FUNCTION_BLOCK FB_FourAxisTrajectory
// 四轴整表轨迹：上位机预检后下发 LREAL 位置点，本块收齐后统一执行。
// 正常流程：0 登记各段 -> 全部下发后 5 统一拼表 -> 0 就绪 -> 10 启动检查 -> 15 首点定位
//           -> 20 开外部给定 -> 30 取点 -> 40 保持末点 -> 60 关闭 -> 70 确认静止 -> 0。
// 异常流程：运动阶段转 50 减速，再经 40/60/70 退出，最后在 90 等待复位。
// 本块每 2 ms 调用一次；使能、点动、回原等基础控制在 FB_AxisControl 中。
// xGroupBusy 占用控制防止两块同时运动，但不能代替设备安全回路。
VAR_INPUT
    xAxesReady : BOOL; // 四轴已使能、回零、静止，供启动和首点定位完成时检查。
    xAbort : BOOL; // 外部联停：许可撤销、撤使能、停止、限位或手动命令冲突。
    nAbortReason : UINT; // MAIN 提供的首个联停原因，0 表示本扫描无联停。
    xAxisFault : BOOL; // 任一轴错误或 NC I/O 反馈无效，拒绝启动或触发联停。
END_VAR
VAR_IN_OUT
    Axes : ARRAY[1..4] OF AXIS_REF; // MAIN 传入的原始轴引用，VAR_IN_OUT 直接操作各 NC 轴接口。
END_VAR
VAR
    // 完整四轴位置表，只由本块分段写入；运行中不再接收上传。
    aPosition : ARRAY[1..4, 0..2099999] OF LREAL; // [轴号, 完整表点号]，所有点号从 0 开始，单位由 NC 配置决定。
    aConfig : ARRAY[1..4] OF ST_AxisConfig; // 启动时锁存参数，首点定位、运行及本次停车使用相同参数。
    aSet : ARRAY[1..4] OF ST_TrajectoryPoint; // 本周期四轴的位置、内部速度和加速度；内部速度用于减速停车。
    aEnable : ARRAY[1..4] OF MC_ExtSetPointGenEnable; // 四个外部给定开启实例；异步执行，等待 NC Enabled 反馈。
    aDisable : ARRAY[1..4] OF MC_ExtSetPointGenDisable; // 四个关闭实例；确认全部退出之前不交回手动。
    aMoveInit : ARRAY[1..4] OF MC_MoveAbsolute; // 四轴各自定位到轨迹首点，全部完成才同步执行位置表。
    aStopInit : ARRAY[1..4] OF MC_Stop; // 外部给定尚未开启时的停车，如取消首点定位。
    rtUpload : R_TRIG; // 本段四轴数据写完后的登记请求上升沿。
    rtAssemble : R_TRIG; // 全部段登记后的独立拼表请求上升沿，不自动启动运动。
    rtClear : R_TRIG; // 清除旧表计数和就绪状态的请求上升沿。
    rtStart : R_TRIG; // 完整位置表就绪后启动轨迹的请求上升沿。
    rtReset : R_TRIG; // 轨迹组故障复位请求上升沿，不复位各 NC 轴故障。
    tmHeartbeat : TON; // 上位机运行心跳超时定时器，启动检查/运动期间 1 秒不变则联停。
    tmEnable : TON; // 四轴外部给定开启阶段超时定时器，限时 5 秒。
    tmMoveInit : TON; // 四轴首点定位阶段超时定时器，限时 60 秒。
    tmExit : TON; // 关闭外部给定及确认退出阶段的超时定时器，限时 5 秒。
    udiLastHeartbeat : UDINT; // 上一扫描上位机运行心跳值，用于检测是否发生变化。
    udiSequence : UDINT; // 当前接收/执行位置表锁存的非零上传序号。
    nCount : UDINT; // 当前整条位置表锁存的单轴总点数，四根轴点数相同。
    nReceived : UDINT; // 已登记的单轴点数，表示段确认进度，不代表已拼入执行表。
    nLoaded : UDINT; // 四轴均已成功拼入执行表的点数。
    nSegment : UDINT; // 当前拼表源段号，从 0 开始，范围 0～20。
    nSegmentPoint : UDINT; // 当前源段内的起始点号，从 0 开始。
    nCopyCount : UDINT; // 本扫描每轴复制点数，受批次、段尾和总表尾三重限制。
    nCopyBytes : UDINT; // 本扫描每轴复制的字节数，等于点数乘 LREAL 大小。
    nSendPoint : UDINT; // 当前轨迹执行取点号，从 0 开始，不是实际到位点号。
    nPrevious : UDINT; // 差分计算前一点索引，首点处夹紧到有效表范围。
    nNext : UDINT; // 差分计算后一点索引，末点处夹紧到有效表范围。
    nHoldCycles : UINT; // 末点静止给定的保持扫描次数，每扫描为 2 ms。
    nStopCycles : UINT; // 减速阶段扫描计数，用于满足该阶段的最少扫描次数。
    nState : UINT; // 轨迹阶段码，数值与上位机监控和故障诊断一致。
    i : INT; // 四轴循环索引，范围 1～4。
    xAllEnabled : BOOL; // 四轴 NC 外部给定均已开启；不是四轴伺服使能汇总。
    xAllDisabled : BOOL; // 四轴外部给定均已关闭，相关开启、关闭和首点停止块均释放 Busy。
    xAllStopped : BOOL; // 四轴 NC 均未处于 Moving 状态；仅为本块此项汇总条件。
    xAllInitDone : BOOL; // 四个首点绝对定位块均输出 Done。
    xMovesIdle : BOOL; // 四个首点定位块均已释放 Busy。
    xEnablePending : BOOL; // 至少一个外部给定开启块仍忙，退出时先等待开启请求结束。
    xFeed : BOOL; // 本扫描需要向四轴发送外部位置给定。
    xValid : BOOL; // 当前轴配置、首点到位或内存复制批次的临时检查结果，每次检查重新赋值。
    xCommandAllowed : BOOL; // 轨迹命令来源为当前有效持有站，且本扫描未发生控制权交接。
    xStopCommand : BOOL; // 当前持有站发出的有效组停止保持命令。
    xUploadRequest : BOOL; // 本扫描获准处理的段登记请求；原始沿已消费后再过滤权限。
    xAssembleRequest : BOOL; // 本扫描获准处理的整表拼接请求。
    xClearRequest : BOOL; // 本扫描获准处理的清表请求。
    xStartRequest : BOOL; // 本扫描获准处理的轨迹启动请求。
    xResetRequest : BOOL; // 本扫描获准处理的轨迹组故障复位请求。
    xNormalStop : BOOL; // 正常人工停止，不作为 1007 故障。
    lrNewVelocity : LREAL; // 当前减速计算的下一扫描速度，单位为 NC 位置单位/秒。
    nBlockAxis : UINT; // 本扫描首个定位/开启块错误的轴，四轴循环结束后统一联停。
    nBlockSource : UINT; // 10=首点定位，11=开启外部给定。
    udiBlockError : UDINT; // 本扫描首个定位/开启块原始错误码，后续轴不能覆盖。
END_VAR
VAR CONSTANT
    // 保留原阶段数值及顺序，供监控和原有区间判断使用。
    cStateIdle : UINT := 0; // 空闲及收段。
    cStateAssemble : UINT := 5; // 拼接已确认的点位段。
    cStateCheckStart : UINT := 10; // 检查轴配置和启动条件。
    cStateMoveToFirstPoint : UINT := 15; // 四轴定位到首点。
    cStateEnableSetpoint : UINT := 20; // 开启外部给定。
    cStateRun : UINT := 30; // 按 2 ms 送点。
    cStateHoldLastPoint : UINT := 40; // 保持末点或停车点。
    cStateDecelerate : UINT := 50; // 减速停车。
    cStateDisableSetpoint : UINT := 60; // 关闭外部给定。
    cStateWaitForStandstill : UINT := 70; // 确认静止并释放组占用。
    cStateFault : UINT := 90; // 等待有效故障复位。
    cDt : LREAL := 0.002; // 单位秒，必须等于 PLC/NC SAF 周期和差分函数周期。
    cMaxPoints : UDINT := 2100000; // 单轴完整表容量，与 aPosition 第二维一致。
    cUploadPoints : UDINT := 100000; // 单轴每段容量，与 GVL_motion.aUpload 第三维一致。
    cCopyPointsPerScan : UDINT := 1024; // 每扫描每轴最多复制 8 KiB；需在目标 PLC 实测任务时间。
END_VAR

// 各 Action 共用本实例变量；运行参数锁存和四轴 MC 实例保持原位。
A01_RequestsAndTimers();
A02_ReadAxisStatus();
A03_ResetAndInterlocks();
// 单一分派：阶段改变后留到下一扫描处理，不能顺序调用三个阶段 Action。
CASE nState OF
cStateIdle, cStateAssemble: A04_ReceiveAndAssemble();
cStateCheckStart, cStateMoveToFirstPoint, cStateEnableSetpoint, cStateRun: A05_PrepareAndRun();
cStateHoldLastPoint, cStateDecelerate, cStateDisableSetpoint, cStateWaitForStandstill: A06_StopAndExit();
END_CASE
// MC 块仍每扫描调用一次，状态发布保持在最后。
A07_CallMotionBlocks();
A08_PublishFeedback();

ACTION A01_RequestsAndTimers:
// 请求、来源站和定时器；写请求沿、诊断首因准备及超时实例。
// 无故障时准备本扫描的诊断位置；故障置位后保持首因，直到有效复位。
IF NOT GVL_motion.xError THEN
    GVL_motion.nFaultAxis := 0;
    GVL_motion.nFaultSource := 0;
    GVL_motion.nFaultState := nState;
    GVL_motion.udiCleanupErrorId := 0;
END_IF
// 1. 上位机操作转为上升沿，防止保持 TRUE 时每扫描重复发起请求。
// 接口顺序：写独立段 -> xUpload 登记 -> 全部段确认 -> xAssemble 统一拼表。
// 原始沿先消费；未授权的保持位不能在以后取得权限时自动变成新请求。
xCommandAllowed := GVL_control.xCanCommand AND NOT GVL_control.xOwnerChanged
    AND (GVL_motion.nCommandStation = GVL_control.nOwner);
xStopCommand := xCommandAllowed AND GVL_motion.xStop;
rtUpload(CLK := GVL_motion.xUpload);
rtAssemble(CLK := GVL_motion.xAssemble);
rtClear(CLK := GVL_motion.xClear);
rtStart(CLK := GVL_motion.xStart);
rtReset(CLK := GVL_motion.xReset);
// Q 是 R_TRIG 的输出，只读取；权限过滤使用独立请求位。
xUploadRequest := rtUpload.Q AND xCommandAllowed;
xAssembleRequest := rtAssemble.Q AND xCommandAllowed;
xClearRequest := rtClear.Q AND xCommandAllowed;
xStartRequest := rtStart.Q AND xCommandAllowed;
xResetRequest := rtReset.Q AND xCommandAllowed;
// 交接或失联使旧表失去启动资格；正在运行时仍走原有联停和退出流程。
IF GVL_control.xOwnerChanged OR NOT GVL_control.xCanCommand THEN
    GVL_motion.xDataReady := FALSE;
    GVL_motion.nUploadStation := 0;
    IF (nState = cStateIdle) OR (nState = cStateAssemble) THEN
        nCount := 0; nReceived := 0; nLoaded := 0; udiSequence := 0; nState := cStateIdle;
    END_IF
END_IF

// 心跳只要变化，TON.IN 就变 FALSE，超时计时复位；连续 1 秒不变则 Q=TRUE。
// 状态 10..40 检查该超时；上传状态 5 不要求心跳，因此可以先上传后开始心跳。
tmHeartbeat(IN := GVL_motion.udiHeartbeat = udiLastHeartbeat, PT := T#1S);
udiLastHeartbeat := GVL_motion.udiHeartbeat;
tmEnable(IN := nState = cStateEnableSetpoint, PT := T#5S);
tmMoveInit(IN := nState = cStateMoveToFirstPoint, PT := T#60S);
tmExit(IN := (nState = cStateDisableSetpoint) OR (nState = cStateWaitForStandstill), PT := T#5S);
IF nState <> cStateDecelerate THEN nStopCycles := 0; END_IF
END_ACTION

ACTION A02_ReadAxisStatus:
// 汇总四轴 NC 状态及 MC 上扫描输出；写六项汇总条件。
// 2. 汇总四轴反馈：AND 从 TRUE 开始，OR 从 FALSE 开始。
// Axis.Status 来自 MAIN 本扫描开头的 ReadStatus。
// 各 MC 块在本块末尾调用，因此这里读到的是它们上一扫描的输出。
xAllEnabled := TRUE;
xAllDisabled := TRUE;
xAllStopped := TRUE;
xAllInitDone := TRUE;
xMovesIdle := TRUE;
xEnablePending := FALSE;
FOR i := 1 TO 4 DO
    xAllEnabled := xAllEnabled AND Axes[i].Status.ExtSetPointGenEnabled;
    // NC 外部给定位为 FALSE 还不够，异步 Enable/Disable 和 Stop.Busy 也要释放。
    // 避免已经交回手动，却仍有上一条异步命令尚未结束。
    xAllDisabled := xAllDisabled AND NOT Axes[i].Status.ExtSetPointGenEnabled
        AND NOT aEnable[i].Busy AND NOT aDisable[i].Busy AND NOT aStopInit[i].Busy;
    xAllStopped := xAllStopped AND NOT Axes[i].Status.Moving;
    xAllInitDone := xAllInitDone AND aMoveInit[i].Done;
    xMovesIdle := xMovesIdle AND NOT aMoveInit[i].Busy;
    xEnablePending := xEnablePending OR aEnable[i].Busy;
END_FOR
END_ACTION

ACTION A03_ResetAndInterlocks:
// 先复位和判断联停，再进入状态机；写首因、停止状态及表资格。
// 复位只清故障；上传完整的位置表保留，新运行仍需使用新的轨迹序号。
// 组复位只清本块故障；各 NC 轴故障仍需通过 Axis1..4.reset 复位。
// 必须已静止、外部给定关闭且相关命令释放，才允许重新进入空闲。
// 未消费序号的上传/启动检查故障可按已确认进度重试；已消费序号需清表并换新序号。
IF xResetRequest AND ((nState = cStateIdle) OR (nState = cStateFault))
    AND xAllStopped AND xAllDisabled AND xMovesIdle THEN
    GVL_motion.xError := FALSE;
    GVL_motion.udiErrorId := 0;
    GVL_motion.nFaultAxis := 0;
    GVL_motion.nFaultSource := 0;
    GVL_motion.nFaultState := 0;
    GVL_motion.udiCleanupErrorId := 0;
    GVL_motion.xDone := FALSE;
    nState := cStateIdle;
END_IF

// 上传阶段不占用轴；启动检查和运动阶段任一轴异常均联停。
// 3. 先判断联停再取点，避免停止条件出现后仍多走一帧。
// 1006=心跳超时，1010=轴错误，1007=停止/联锁/冲突/外部给定意外退出。
// 状态 10 尚未发运动命令，可直接进 90；其他阶段先进 50 减速退出。
// 故障置位后不重复把状态 40 拉回 50，保证末点保持和退出可以完成。
IF (nState >= cStateCheckStart) AND (nState <= cStateHoldLastPoint) AND NOT GVL_motion.xError THEN
    IF xAxisFault OR xAbort OR tmHeartbeat.Q
        OR ((nState >= cStateRun) AND NOT xAllEnabled) THEN
        GVL_motion.xError := TRUE;
        IF tmHeartbeat.Q THEN
            GVL_motion.udiErrorId := 1006;
            GVL_motion.nFaultSource := 7;
        ELSIF xAxisFault THEN
            GVL_motion.udiErrorId := 1010;
            GVL_motion.nFaultSource := 8;
            FOR i := 1 TO 4 DO
                IF Axes[i].Status.Error OR Axes[i].Status.IoDataInvalid
                    OR ((i = 1) AND GVL_axis.Axis1.xError) OR ((i = 2) AND GVL_axis.Axis2.xError)
                    OR ((i = 3) AND GVL_axis.Axis3.xError) OR ((i = 4) AND GVL_axis.Axis4.xError) THEN
                    GVL_motion.nFaultAxis := INT_TO_UINT(i); EXIT;
                END_IF
            END_FOR
        ELSE
            GVL_motion.udiErrorId := 1007;
            IF xAbort THEN GVL_motion.nFaultSource := nAbortReason;
            ELSE GVL_motion.nFaultSource := 9;
            END_IF
        END_IF
        IF nState = cStateCheckStart THEN nState := cStateFault; ELSE nState := cStateDecelerate; END_IF
    END_IF
END_IF

// 人工停止：取消收段/拼表/启动检查，运动阶段从当前给定减速；不人为生成故障。
IF xStopCommand AND NOT GVL_motion.xError THEN
    xNormalStop := TRUE;
    GVL_motion.xDataReady := FALSE;
    GVL_motion.xDone := FALSE;
    IF (nState = cStateIdle) OR (nState = cStateAssemble) OR (nState = cStateCheckStart) THEN
        nCount := 0; nReceived := 0; nLoaded := 0; udiSequence := 0; nState := cStateIdle;
        GVL_motion.xStopped := xAllStopped AND xAllDisabled AND xMovesIdle;
    ELSIF (nState = cStateMoveToFirstPoint) OR (nState = cStateEnableSetpoint) OR (nState = cStateRun) THEN
        nStopCycles := 0;
        nState := cStateDecelerate;
    END_IF
END_IF
END_ACTION

ACTION A04_ReceiveAndAssemble:
// 状态 0/5：收段、清表、拼表和启动请求登记；不推进运动点。
CASE nState OF

cStateIdle: // 空闲：先接收所有独立段，再统一拼表；拼接完成后才允许启动。
    // 清表只清计数和就绪状态，不遍历清零约 134.4 MB 的接收区和执行表。
    // 新轨迹必须从偏移 0 连续覆盖所有有效点，旧数据不会在未收齐时被执行。
    // 同扫描多个请求的优先级为 Clear -> Upload -> Assemble -> Start。
    IF xStopCommand THEN
        // 停止保持期间不接受同扫描上传/拼接/启动请求。
    ELSIF xClearRequest AND xAllDisabled AND xMovesIdle THEN
        xNormalStop := FALSE;
        GVL_motion.xStopped := FALSE;
        GVL_motion.nUploadStation := GVL_control.nOwner;
        nCount := 0;
        nReceived := 0;
        nLoaded := 0;
        udiSequence := 0;
        GVL_motion.xDataReady := FALSE;
        GVL_motion.xDone := FALSE;
    ELSIF xUploadRequest AND NOT GVL_motion.xError THEN
        // 只登记写完的独立段，此处不复制任何位置点。
        // 连续偏移及固定段长共同避免漏段、重复段和错段；先检查范围再做 UDINT 减法。
        IF (GVL_motion.nPointCount < 4) OR (GVL_motion.nPointCount > cMaxPoints)
            OR (GVL_motion.nSampleTimeUs <> 2000) OR (GVL_motion.udiUploadSequence = 0)
            OR (GVL_motion.udiUploadSequence = GVL_motion.udiAcceptedSequence)
            OR (GVL_motion.nUploadCount = 0) OR (GVL_motion.nUploadCount > cUploadPoints)
            OR (GVL_motion.nUploadOffset <> nReceived) THEN
            GVL_motion.udiErrorId := 1001;
            GVL_motion.nFaultSource := 17;
        ELSIF nReceived > GVL_motion.nPointCount THEN
            GVL_motion.udiErrorId := 1001;
            GVL_motion.nFaultSource := 17;
        ELSIF GVL_motion.nUploadCount <> MIN(cUploadPoints, GVL_motion.nPointCount - nReceived) THEN
            GVL_motion.udiErrorId := 1001;
            GVL_motion.nFaultSource := 17;
        ELSIF (nReceived <> 0) AND ((GVL_motion.nPointCount <> nCount)
            OR (GVL_motion.udiUploadSequence <> udiSequence)) THEN
            GVL_motion.udiErrorId := 1001;
            GVL_motion.nFaultSource := 17;
        ELSE
            // 接收确认只表示 PC 已声明本段四轴写完；ADS 数据仍须由 PC 遵守只写一次的约定。
            GVL_motion.nUploadStation := GVL_control.nOwner;
            GVL_motion.xStopped := FALSE;
            xNormalStop := FALSE;
            nCount := GVL_motion.nPointCount;
            udiSequence := GVL_motion.udiUploadSequence;
            nReceived := nReceived + GVL_motion.nUploadCount;
            GVL_motion.xDataReady := FALSE;
        END_IF
        IF GVL_motion.udiErrorId <> 0 THEN
            GVL_motion.xError := TRUE;
            nState := cStateFault;
        END_IF
    ELSIF xAssembleRequest AND NOT GVL_motion.xError THEN
        // 必须收到全部段的确认和独立的完成请求，不能因最后一段到齐就自动拼表或启动。
        IF (nCount < 4) OR (nReceived <> nCount) OR (udiSequence = 0)
            OR (udiSequence = GVL_motion.udiAcceptedSequence)
            OR (GVL_motion.nPointCount <> nCount) OR (GVL_motion.nSampleTimeUs <> 2000)
            OR (GVL_motion.udiUploadSequence <> udiSequence) THEN
            GVL_motion.xError := TRUE;
            GVL_motion.udiErrorId := 1001;
            GVL_motion.nFaultSource := 17;
            nState := cStateFault;
        ELSE
            nLoaded := 0;
            GVL_motion.xDataReady := FALSE;
            GVL_motion.xDone := FALSE;
            nState := cStateAssemble;
        END_IF
    ELSIF xStartRequest AND NOT GVL_motion.xError THEN
        GVL_motion.xDone := FALSE;
        GVL_motion.nCurrentPoint := 0;
        // 点位数值由上位机预检；上传完整只代表表已收齐，不代表轴已到首点。
        // 禁止重放已消费序号，避免旧启动命令重复执行轨迹。
        IF NOT GVL_motion.xDataReady OR (GVL_motion.nUploadStation <> GVL_control.nOwner) OR (nLoaded <> nCount) OR (nCount < 4)
            OR (udiSequence = GVL_motion.udiAcceptedSequence)
            OR (GVL_motion.nPointCount <> nCount) OR (GVL_motion.nSampleTimeUs <> 2000)
            OR (GVL_motion.udiUploadSequence <> udiSequence) THEN
            GVL_motion.udiErrorId := 1001;
            GVL_motion.nFaultSource := 17;
        ELSIF NOT xAxesReady OR NOT xAllDisabled OR NOT xMovesIdle
            OR xAbort OR GVL_motion.xStop OR xAxisFault OR tmHeartbeat.Q THEN
            GVL_motion.udiErrorId := 1004;
            GVL_motion.nFaultSource := 16;
        ELSE
            // 锁存本次运行参数；配置仅应在轴静止且轨迹空闲时修改。
            // 状态 10 仅检查轴配置和就绪，随后进入首点定位。
            aConfig := GVL_motion.aConfig;
            nState := cStateCheckStart;
        END_IF
        IF GVL_motion.udiErrorId <> 0 THEN
            GVL_motion.xError := TRUE;
            nState := cStateFault;
        END_IF
    END_IF

cStateAssemble: // 全部段下发后才进入这里，按段号拼入四轴连续表，PC 不得再改接收区。
    IF (GVL_motion.nPointCount <> nCount) OR (GVL_motion.udiUploadSequence <> udiSequence)
        OR (GVL_motion.nSampleTimeUs <> 2000) OR xUploadRequest OR xClearRequest OR xAssembleRequest THEN
        // 元数据或请求冲突使本次拼接失效；复位后重新 xAssemble，从第 0 点重拼。
        GVL_motion.xError := TRUE;
        GVL_motion.udiErrorId := 1001;
        GVL_motion.nFaultSource := 17;
        nState := cStateFault;
    ELSE
        nSegment := nLoaded / cUploadPoints;
        nSegmentPoint := nLoaded MOD cUploadPoints;
        // 同时限制本拍工作量、剩余总点数和当前段剩余量，短末段也不会越界或串轴。
        nCopyCount := MIN(cCopyPointsPerScan, MIN(nCount - nLoaded, cUploadPoints - nSegmentPoint));
        nCopyBytes := nCopyCount * SIZEOF(aPosition[1, 0]);
        xValid := TRUE;
        FOR i := 1 TO 4 DO
            // 每轴只做一次有界内存复制；源/目标独立，地址每扫描现取，不缓存指针。
            IF MEMCPY(destAddr := ADR(aPosition[i, nLoaded]),
                srcAddr := ADR(GVL_motion.aUpload[nSegment, i, nSegmentPoint]), n := nCopyBytes) <> nCopyBytes THEN
                xValid := FALSE;
            END_IF
        END_FOR
        IF NOT xValid THEN
            GVL_motion.xError := TRUE;
            GVL_motion.udiErrorId := 1012;
            GVL_motion.nFaultSource := 18;
            nState := cStateFault;
        ELSE
            // 四轴本批全部复制成功才推进；最后一批完成后才发布整表就绪。
            nLoaded := nLoaded + nCopyCount;
            IF nLoaded = nCount THEN GVL_motion.xDataReady := TRUE; nState := cStateIdle; END_IF
        END_IF
    END_IF

END_CASE
END_ACTION

ACTION A05_PrepareAndRun:
// 状态 10/15/20/30：检查配置、首点、开启、同步取点；一次只执行当前分支。
CASE nState OF

cStateCheckStart: // 单扫描检查配置与轴就绪；整表数值已由上位机在发送前预检。
    // PLC 不再遍历点位表；保留锁存配置检查，供首点定位、运行及停车使用。
    FOR i := 1 TO 4 DO
        xValid := F_AxisConfigValid(aConfig[i])
            AND (aConfig[i].lrStartTolerance > 0) AND (aConfig[i].lrStartTolerance < 1.0E6)
            AND (aConfig[i].lrInitVelocity > 0) AND (aConfig[i].lrInitVelocity <= aConfig[i].lrMaxVelocity);
        IF NOT xValid THEN
            GVL_motion.udiErrorId := 1002;
            GVL_motion.nFaultAxis := INT_TO_UINT(i);
            GVL_motion.nFaultSource := 15;
            EXIT;
        END_IF
    END_FOR
    IF GVL_motion.udiErrorId <> 0 THEN
        GVL_motion.xError := TRUE;
        nState := cStateFault;
    ELSIF NOT xAxesReady THEN
        GVL_motion.xError := TRUE;
        GVL_motion.udiErrorId := 1004;
        GVL_motion.nFaultSource := 16;
        nState := cStateFault;
    ELSE
        FOR i := 1 TO 4 DO
            aSet[i].lrPosition := aPosition[i, 0];
            aSet[i].lrVelocity := 0;
            aSet[i].lrAcceleration := 0;
        END_FOR
        // 启动检查通过后消费序号；首点定位即使失败，也须换新序号重发。
        GVL_motion.udiAcceptedSequence := udiSequence;
        nSendPoint := 0;
        nState := cStateMoveToFirstPoint;
    END_IF

cStateMoveToFirstPoint: // 参考旧工程 move_init：四轴各自定位到首点，全部完成才激活外部给定。
    // 状态 15 让下方 MoveAbsolute.Execute 产生上升沿，速度用 lrInitVelocity。
    // 四轴定位各自规划，到位时间可不同；全部 Done 并检查实际/设定位置偏差后才同步取点。
    // 超过 60 秒报 1011；停止定位需要 MC_Stop，不能只把 MoveAbsolute.Execute 清零。
    IF tmMoveInit.Q THEN
        GVL_motion.xError := TRUE;
        GVL_motion.udiErrorId := 1011;
        GVL_motion.nFaultSource := 19;
        nState := cStateDecelerate;
    ELSIF xAllInitDone AND xAxesReady THEN
        xValid := TRUE;
        FOR i := 1 TO 4 DO
            IF NOT ((ABS(Axes[i].NcToPlc.ActPos - aPosition[i, 0]) <= aConfig[i].lrStartTolerance)
                AND (ABS(Axes[i].NcToPlc.SetPos - aPosition[i, 0]) <= aConfig[i].lrStartTolerance)) THEN
                IF xValid THEN GVL_motion.nFaultAxis := INT_TO_UINT(i); END_IF
                xValid := FALSE;
            END_IF
        END_FOR
        IF xValid THEN nState := cStateEnableSetpoint;
        ELSE
            GVL_motion.xError := TRUE;
            GVL_motion.udiErrorId := 1004;
            GVL_motion.nFaultSource := 16;
            nState := cStateDecelerate;
        END_IF
    END_IF

cStateEnableSetpoint: // 四轴激活过程中持续送静止首点，共同确认后才推进点号。
    // 状态 20 发起异步外部给定开启请求；等待期间仍送静止首点，不推进点号。
    // 用四根轴的 ExtSetPointGenEnabled 汇总确认，而不是只等其中某个 Enable.Done。
    IF tmEnable.Q THEN
        GVL_motion.xError := TRUE;
        GVL_motion.udiErrorId := 1008;
        GVL_motion.nFaultSource := 20;
        nState := cStateDecelerate;
    ELSIF xAllEnabled THEN nState := cStateRun;
    END_IF

cStateRun: // 位置取点方式与参考工程相同，四轴共用 nSendPoint。
    // 四轴都读取同一个 nSendPoint，每扫描只在四轴循环后推进一次点号。
    // 共享点号保证设定值在同一扫描更新，实际跟随误差由各轴 NC/驱动器反馈决定。
    // 相邻位置点转换为速度/加速度，上位机无需额外下发这两个数组。
    nPrevious := nSendPoint;
    IF nSendPoint > 0 THEN nPrevious := nSendPoint - 1; END_IF
    nNext := MIN(nSendPoint + 1, nCount - 1);
    FOR i := 1 TO 4 DO
        aSet[i] := F_TrajectoryPoint(lrPrevious := aPosition[i, nPrevious],
            lrCurrent := aPosition[i, nSendPoint], lrNext := aPosition[i, nNext],
            xEndpoint := (nSendPoint = 0) OR (nSendPoint = nCount - 1));
    END_FOR
    // 反馈的是本扫描准备送出的点号；递增 nSendPoint 只影响下一次状态 30。
    // 本扫描末尾的 Feed 仍发送已经保存在 aSet 中的当前点。
    GVL_motion.nCurrentPoint := nSendPoint;
    IF nSendPoint = nCount - 1 THEN nHoldCycles := 0; nState := cStateHoldLastPoint;
    ELSE nSendPoint := nSendPoint + 1;
    END_IF

END_CASE
END_ACTION

ACTION A06_StopAndExit:
// 状态 40/50/60/70：保持、减速、关闭和退出；故障 90 等待有效复位。
CASE nState OF

cStateHoldLastPoint: // 末点静止给定保持两个周期，随后关闭外部给定，不强制跳回零位。
    // 正常末点和减速终点都到这里；设定速度已经为 0。
    // 静止点多保持两拍，给 NC 消费最后给定留出时间，再发关闭命令。
    FOR i := 1 TO 4 DO aSet[i].lrAcceleration := 0; END_FOR
    nHoldCycles := nHoldCycles + 1;
    IF nHoldCycles >= 2 THEN nState := cStateDisableSetpoint; END_IF

cStateDecelerate: // 外部轨迹按最后的设定速度减速；首点定位由下方 MC_Stop 停车。
    // 至少经过一次 Stop 调用再退出，覆盖定位请求刚被取消但实际轴仍在运动的情况。
    IF nStopCycles < 2 THEN nStopCycles := nStopCycles + 1; END_IF
    xValid := TRUE;
    FOR i := 1 TO 4 DO
        // 正速度逐步降到 0，负速度逐步升到 0，MAX/MIN 防止跨零反向。
        // 各轴停车减速度独立，停车时刻/距离可能不同，不维持四轴路径比例。
        IF aSet[i].lrVelocity > 0 THEN
            lrNewVelocity := MAX(0, aSet[i].lrVelocity - aConfig[i].lrStopDeceleration * cDt);
        ELSE lrNewVelocity := MIN(0, aSet[i].lrVelocity + aConfig[i].lrStopDeceleration * cDt);
        END_IF
        // 位置用梯形积分：pNew=pOld+(vOld+vNew)/2*dt；加速度=(vNew-vOld)/dt。
        // 从最后给定连续减速，不跳到轨迹末点；本实现未加入 jerk 平滑。
        aSet[i].lrPosition := aSet[i].lrPosition + (aSet[i].lrVelocity + lrNewVelocity) * 0.5 * cDt;
        aSet[i].lrAcceleration := (lrNewVelocity - aSet[i].lrVelocity) / cDt;
        aSet[i].lrVelocity := lrNewVelocity;
        xValid := xValid AND (lrNewVelocity = 0);
    END_FOR
    // 外部给定未退出时 NC 的 Moving 可能仍有效；先结束设定减速，再退出并等待实际静止。
    IF xValid AND xMovesIdle AND (nStopCycles >= 2) THEN nHoldCycles := 0; nState := cStateHoldLastPoint; END_IF

cStateDisableSetpoint: // 等待异步 Enable 结束后再 Disable，防止迟到的 Enable 再次打开轴。
    // xAllDisabled 同时检查 NC 标志和 MC.Busy；关闭失败时保持此状态占用。
    // 复位沿可使下方 Disable 暂时撤请求，下一拍重新产生上升沿进行重试。
    IF xAllDisabled THEN nState := cStateWaitForStandstill; END_IF

// 状态 70：关闭命令完成后，再等实际轴静止及定位命令释放。
// 正常结束才置 xDone；发生过联停/故障则转 90，避免误报正常完成。
// 状态 90 没有 CASE 动作，保留故障，等待上方符合条件的复位沿。
cStateWaitForStandstill:
    IF xAllStopped AND xAllDisabled AND xMovesIdle THEN
        IF GVL_motion.xError THEN nState := cStateFault;
        ELSIF xNormalStop THEN GVL_motion.xStopped := TRUE; nState := cStateIdle;
        ELSE GVL_motion.xDone := TRUE; nState := cStateIdle;
        END_IF
    END_IF

END_CASE
END_ACTION

ACTION A07_CallMotionBlocks:
// 每扫描调用四轴 MC 实例，循环结束统一处理错误；写 MC 输出及清理错误。
// 功能块每周期调用；禁止在四轴循环中途改变公共状态。
// 5. 外部给定实际入口：下面的 Feed、Enable、Disable。
// 状态 20 等开启、30 取点、40 保持、50 减速、60 等关闭，都需要持续更新给定。
// 状态 15 用内部 MoveAbsolute 定位，不执行外部轨迹运动。
// 关闭请求发出后仍送静止点，直到 NC 确认外部给定已关闭。
xFeed := (nState >= cStateEnableSetpoint) AND (nState <= cStateDisableSetpoint);
udiBlockError := 0;
nBlockAxis := 0;
nBlockSource := 0;
FOR i := 1 TO 4 DO
    // A. 首点定位：每轴实例保存自己的 Busy/Done/Error，每扫描都要继续调用。
    // Execute 下降沿不等于立即停止，取消时由下面 MC_Stop 完成停车。
    aMoveInit[i](Axis := Axes[i], Execute := nState = cStateMoveToFirstPoint,
        Position := aPosition[i, 0], Velocity := aConfig[i].lrInitVelocity,
        Acceleration := aConfig[i].lrMaxAcceleration, Deceleration := aConfig[i].lrStopDeceleration);
    // B. 尚未开启外部给定的轴使用 MC_Stop；已开启的轴由状态 50 生成减速给定。
    // 避免外部给定有效时同时用 Stop 和 Feed 争用同一根轴。
    aStopInit[i](Axis := Axes[i], Execute := (nState = cStateDecelerate) AND NOT Axes[i].Status.ExtSetPointGenEnabled,
        Deceleration := aConfig[i].lrStopDeceleration);
    IF xFeed THEN
        // C. 送绝对位置，按确认的调用方式固定速度 0、加速度 2000。
        // Direction 固定为 1，使 NC 在运行、反向和末点保持期间持续采纳位置。
        // PLC 内部仍用 aSet 的速度计算减速停车点位。
        // 该函数返回值不代表本点执行完成，不能用它控制 nSendPoint 递增。
        MC_ExtSetPointGenFeed(Axis := Axes[i],
                            Position := aSet[i].lrPosition,
                            Velocity := 0.0,
                            Acceleration := 2000.0,
                            Direction := 1);
    END_IF
    // D. 开启外部给定：状态 20 的 Execute 上升沿发起异步命令。
    // PositionType=ABSOLUTE；Position 传末点用于目标位置监控，不是让轴立即跑到末点。
    // 轴每拍具体走到哪里，由 Feed.Position 决定；首点定位已由 A 完成。
    // MAX(nCount,1)-1 保证空闲时 nCount=0 也只访问第 0 点，不发生 UDINT 下溢。
                aEnable[i](Axis := Axes[i],
                Execute := nState = cStateEnableSetpoint,
                Position := aPosition[i, MAX(nCount, 1) - 1],
                PositionType := POSITIONTYPE_ABSOLUTE);
    // E. 关闭外部给定：状态 60 请求，先等所有开启请求 Busy 结束。
    // xResetRequest 暂时撤销 Execute，下一拍恢复形成新上升沿，供关闭失败后重试。
    // 确认关闭后还需经过状态 70，才把轴交回基础手动控制。
    aDisable[i](Axis := Axes[i],
                Execute := (nState = cStateDisableSetpoint) AND NOT xEnablePending AND NOT xResetRequest);

    // 四轴仍执行同一阶段；只登记最先出错的轴，循环结束后统一改变状态。
    IF nBlockAxis = 0 THEN
        IF aMoveInit[i].Error AND (nState = cStateMoveToFirstPoint) THEN
            udiBlockError := aMoveInit[i].ErrorID; nBlockAxis := INT_TO_UINT(i); nBlockSource := 10;
        ELSIF aEnable[i].Error AND (nState = cStateEnableSetpoint) THEN
            udiBlockError := aEnable[i].ErrorID; nBlockAxis := INT_TO_UINT(i); nBlockSource := 11;
        END_IF
    END_IF
    // 清理错误单独保存；此前已有故障时不能覆盖原始错误号和来源。
    IF ((aStopInit[i].Error AND (nState = cStateDecelerate)) OR (aDisable[i].Error AND (nState = cStateDisableSetpoint)))
        AND (GVL_motion.udiCleanupErrorId = 0) THEN
        IF nState = cStateDecelerate THEN GVL_motion.udiCleanupErrorId := aStopInit[i].ErrorID;
        ELSE GVL_motion.udiCleanupErrorId := aDisable[i].ErrorID;
        END_IF
        IF GVL_motion.udiCleanupErrorId = 0 THEN GVL_motion.udiCleanupErrorId := 1009; END_IF
        IF NOT GVL_motion.xError THEN
            GVL_motion.udiErrorId := GVL_motion.udiCleanupErrorId;
            GVL_motion.nFaultAxis := INT_TO_UINT(i);
            IF nState = cStateDecelerate THEN GVL_motion.nFaultSource := 12;
            ELSE GVL_motion.nFaultSource := 13;
            END_IF
            GVL_motion.nFaultState := nState;
            GVL_motion.xError := TRUE;
        END_IF
    END_IF
END_FOR
IF nBlockAxis <> 0 THEN
    IF NOT GVL_motion.xError THEN
        GVL_motion.udiErrorId := udiBlockError;
        IF udiBlockError = 0 THEN GVL_motion.udiErrorId := 1010; END_IF
        GVL_motion.nFaultAxis := nBlockAxis;
        GVL_motion.nFaultSource := nBlockSource;
        GVL_motion.nFaultState := nState;
        GVL_motion.xError := TRUE;
    END_IF
    nState := cStateDecelerate;
END_IF
// 退出超时只报错，不强行清 Busy 或改回空闲，防止仍被占用的轴接受新运动。
IF tmExit.Q AND ((nState = cStateDisableSetpoint) OR (nState = cStateWaitForStandstill)) THEN
    IF GVL_motion.udiCleanupErrorId = 0 THEN GVL_motion.udiCleanupErrorId := 1009; END_IF
    IF NOT GVL_motion.xError THEN
        GVL_motion.udiErrorId := 1009;
        GVL_motion.nFaultSource := 14;
        GVL_motion.nFaultState := nState;
        GVL_motion.xError := TRUE;
    END_IF
END_IF
END_ACTION

ACTION A08_PublishFeedback:
// 最后发布接收、拼接、状态和占用反馈；不写运动命令。
// 6. 已接收和已拼接分开发布；只有 xDataReady 才表示完整表可进入启动检查。
GVL_motion.nReceivedCount := nReceived;
GVL_motion.udiReceivedSequence := udiSequence;
GVL_motion.nLoadedCount := nLoaded;
GVL_motion.nState := nState;
GVL_motion.xUploadBusy := nState = cStateAssemble;
GVL_motion.xBusy := (nState >= cStateCheckStart) AND (nState <= cStateWaitForStandstill);
GVL_motion.xRunning := nState = cStateRun;
END_ACTION

END_FUNCTION_BLOCK

(* stored: Version 1.1.0.1
   POU FB_FourAxisTrajectory: Id {f339b171-2adc-4ce0-8fc1-1403fdabbc80}, SpecialFunc None
   Action A01_RequestsAndTimers: Id {332b3d73-5f1e-53b4-bfd7-3498fa26ebc9}
   Action A02_ReadAxisStatus: Id {3309f391-5387-5da0-bdd1-bf0a7f5a76a5}
   Action A03_ResetAndInterlocks: Id {6e12063d-0d55-579e-87d7-4b0052990f27}
   Action A04_ReceiveAndAssemble: Id {d38f3d56-ae53-5674-96cb-a2428028aced}
   Action A05_PrepareAndRun: Id {3069ae07-2eca-5a5e-ab04-53abc58ef09f}
   Action A06_StopAndExit: Id {d1256174-2d27-54a4-9857-8a726236adaa}
   Action A07_CallMotionBlocks: Id {385add14-f0d7-5c01-a475-a0408dc09db6}
   Action A08_PublishFeedback: Id {57401618-0d32-59ac-acf9-fa630b378184} *)
